{region 'Documentation'}
(*!
<summary>Copies a small fixed child view and records actual-index access by the helper.</summary>
<description>
Initialize reads real bounds from the fixture's selected fixed array and copies only
its registered prefix. The copy is intentional test-double storage, not a production
registry or retained array pointer. GetChild translates the original index without
calling a child. Invalid access and trace overflow remain observable.
</description>
*)
{endregion}
FUNCTION_BLOCK OrchestrationCollectionDouble IMPLEMENTS I_OrchestratableCollection
VAR
    FChildren : ARRAY[1..ChildCapacity] OF I_Orchestratable;
    FLowerBound : DINT;
    FUpperBound : DINT;
    FCount : UINT;
    FReadIndices : ARRAY[1..ReadCapacity] OF DINT;
    FReadCount : UINT;
    FInvalidAccess : BOOL;
    FTraceOverflow : BOOL;
END_VAR
VAR CONSTANT
    ChildCapacity : UINT := 3;
    ReadCapacity : UINT := 512;
END_VAR

{region 'Documentation'}
(*!
<summary>Actual input-array lower bound.</summary>
*)
{endregion}
{attribute 'monitoring' := 'call'}
PROPERTY PUBLIC ChildArrayLowerBound : DINT //! Actual input-array lower bound.
GET
ChildArrayLowerBound := FLowerBound;
END_GET
END_PROPERTY

{region 'Documentation'}
(*!
<summary>Actual input-array capacity upper bound.</summary>
*)
{endregion}
{attribute 'monitoring' := 'call'}
PROPERTY PUBLIC ChildArrayUpperBound : DINT //! Actual input-array capacity upper bound.
GET
ChildArrayUpperBound := FUpperBound;
END_GET
END_PROPERTY

{region 'Documentation'}
(*!
<summary>Number of occupied entries.</summary>
*)
{endregion}
{attribute 'monitoring' := 'call'}
PROPERTY PUBLIC ChildCount : UINT //! Number of occupied entries.
GET
ChildCount := FCount;
END_GET
END_PROPERTY

{region 'Documentation'}
(*!
<summary>Records the original array index and returns only registered entries; never invokes a child.</summary>
*)
{endregion}
METHOD PUBLIC GetChild : I_Orchestratable //! Copied child interface at the original occupied index; zero and a latched InvalidAccess for an invalid index.
VAR_INPUT
    Index : DINT; //! Original array index to record and resolve within the occupied prefix.
END_VAR
VAR
    Position : LINT;
END_VAR
GetChild := 0;
IF FReadCount < ReadCapacity THEN
    FReadCount := FReadCount + 1;
    FReadIndices[FReadCount] := Index;
ELSE
    FTraceOverflow := TRUE;
END_IF;

Position := DINT_TO_LINT(Index) - DINT_TO_LINT(FLowerBound) + 1;
IF (Position < 1) OR (Position > UINT_TO_LINT(FCount)) THEN
    FInvalidAccess := TRUE;
    RETURN;
END_IF;
GetChild := FChildren[LINT_TO_UINT(Position)];
END_METHOD

{region 'Documentation'}
(*!
<summary>Copies the fixed registered prefix and clears access evidence without retaining addresses.</summary>
*)
{endregion}
METHOD PUBLIC Initialize : BOOL //! TRUE after copying a valid nonzero occupied prefix; FALSE leaves ChildCount zero.
VAR_INPUT
    Count : UINT; //! Occupied prefix length in 1..ChildCapacity; it must fit the supplied array.
END_VAR
VAR_IN_OUT
    Children : ARRAY[*] OF I_Orchestratable; //! Borrowed array whose occupied interface prefix is copied; keep the referenced children alive.
END_VAR
VAR
    Position : UINT;
    ArrayIndex : DINT;
END_VAR
Initialize := FALSE;
FCount := 0;
FLowerBound := LOWER_BOUND(Children, 1);
FUpperBound := UPPER_BOUND(Children, 1);
FReadCount := 0;
FInvalidAccess := FALSE;
FTraceOverflow := FALSE;
FOR Position := 1 TO ChildCapacity DO
    FChildren[Position] := 0;
END_FOR;
FOR Position := 1 TO ReadCapacity DO
    FReadIndices[Position] := 0;
END_FOR;
IF (Count = 0) OR (Count > ChildCapacity)
    OR (DINT_TO_LINT(FLowerBound) + UINT_TO_LINT(Count) - 1 > DINT_TO_LINT(FUpperBound)) THEN
    RETURN;
END_IF;

FOR Position := 1 TO Count DO
    ArrayIndex := FLowerBound + UINT_TO_DINT(Position) - 1;
    IF Children[ArrayIndex] = 0 THEN
        RETURN;
    END_IF;
    FChildren[Position] := Children[ArrayIndex];
END_FOR;
FCount := Count;
Initialize := TRUE;
END_METHOD

{region 'Documentation'}
(*!
<summary>Latched access outside the registered range.</summary>
*)
{endregion}
{attribute 'monitoring' := 'call'}
PROPERTY PUBLIC InvalidAccess : BOOL //! Latched access outside the registered range.
GET
InvalidAccess := FInvalidAccess;
END_GET
END_PROPERTY

{region 'Documentation'}
(*!
<summary>Number of retained index-access observations.</summary>
*)
{endregion}
{attribute 'monitoring' := 'call'}
PROPERTY PUBLIC ReadCount : UINT //! Number of retained index-access observations.
GET
ReadCount := FReadCount;
END_GET
END_PROPERTY

{region 'Documentation'}
(*!
<summary>Whether the bounded index trace was exhausted.</summary>
*)
{endregion}
{attribute 'monitoring' := 'call'}
PROPERTY PUBLIC TraceOverflow : BOOL //! Whether the bounded index trace was exhausted.
GET
TraceOverflow := FTraceOverflow;
END_GET
END_PROPERTY

END_FUNCTION_BLOCK

(* stored: Version 1.1.0.1
   POU OrchestrationCollectionDouble: Id {0f2e9bb6-f6ba-479c-9a8d-c7556a88b772}, SpecialFunc None
   Property ChildArrayLowerBound: Id {f5e4eb33-88f1-4926-9a6c-1ca1453ce1da}
   Get Get: Id {53075e1e-f107-49e3-985e-19efd0d8b37f}
   Property ChildArrayUpperBound: Id {dc4a9d96-a7aa-4f55-bfb2-86faed04f6f4}
   Get Get: Id {897d1ad8-a809-4778-a5e2-3369250be454}
   Property ChildCount: Id {15950828-9c47-46f0-807d-bbca17d5915b}
   Get Get: Id {9ce7ce1c-afb8-40a2-b511-675cd881fcc3}
   Method GetChild: Id {53a4bdbb-b9fd-4e0b-b7bf-0af8008a3ebb}
   Method Initialize: Id {96d3e0af-aab3-4fdf-999b-62be6b66f807}
   Property InvalidAccess: Id {37afb7e1-0196-4eb6-a5e2-f807522399bc}
   Get Get: Id {6dd2fae8-4911-4bad-9350-bc37bfd0a475}
   Property ReadCount: Id {8a615a60-4867-4a5d-9d10-4f357d1fc258}
   Get Get: Id {c361f4f2-a8fb-4dea-a5fb-f560660b95db}
   Property TraceOverflow: Id {fdb74941-d67f-4bb1-9ce7-0c7774dbf895}
   Get Get: Id {2e6b2f17-a219-4a72-8516-c466a3e04b9d} *)
